(* IEC 61131-3 sources: OpenPlc_Lezioni/Blocchi_PorteLogiche/build, 2 files *)

(* ---- plc.st ---- *)
TYPE
  LOGLEVEL : (CRITICAL, WARNING, INFO, DEBUG) := INFO;
END_TYPE

FUNCTION_BLOCK LOGGER
  VAR_INPUT
    TRIG : BOOL;
    MSG : STRING;
    LEVEL : LOGLEVEL := INFO;
  END_VAR
  VAR
    TRIG0 : BOOL;
  END_VAR

  IF TRIG AND NOT TRIG0 THEN
  {{
   LogMessage(GetFbVar(LEVEL),(char*)GetFbVar(MSG, .body),GetFbVar(MSG, .len));
  }}
  END_IF;
  TRIG0:=TRIG;
END_FUNCTION_BLOCK

PROGRAM program0
  VAR
    P1 : BOOL;
    P2 : BOOL;
    P3 : BOOL;
    P4 : BOOL;
    P5 : BOOL;
    P6 : BOOL;
    P7 : BOOL;
    LED1 : BOOL;
    LED2 : BOOL;
    LED3 : BOOL;
    LED4 : BOOL;
    _TMP_AND1_OUT : BOOL;
    _TMP_OR2_OUT : BOOL;
    _TMP_AND10_OUT : BOOL;
    _TMP_NOT18_OUT : BOOL;
  END_VAR

  _TMP_AND1_OUT := AND(P1, P2);
  LED1 := _TMP_AND1_OUT;
  _TMP_OR2_OUT := OR(P3, P4);
  LED2 := _TMP_OR2_OUT;
  _TMP_AND10_OUT := AND(P5, P6);
  LED2 := _TMP_AND10_OUT;
  _TMP_NOT18_OUT := NOT(P7);
  LED4 := _TMP_NOT18_OUT;
END_PROGRAM

CONFIGURATION Config0

  RESOURCE Res0 ON PLC
    TASK task0(INTERVAL := T#20ms,PRIORITY := 0);
    PROGRAM instance0 WITH task0 : program0;
  END_RESOURCE
END_CONFIGURATION

(* ---- generated_plc.st ---- *)
PROGRAM program0
  VAR
    P1 : BOOL;
    P2 : BOOL;
    P3 : BOOL;
    P4 : BOOL;
    P5 : BOOL;
    P6 : BOOL;
    P7 : BOOL;
    LED1 : BOOL;
    LED2 : BOOL;
    LED3 : BOOL;
    LED4 : BOOL;
    _TMP_AND1_OUT : BOOL;
    _TMP_OR2_OUT : BOOL;
    _TMP_AND10_OUT : BOOL;
    _TMP_NOT18_OUT : BOOL;
  END_VAR

  _TMP_AND1_OUT := AND(P1, P2);
  LED1 := _TMP_AND1_OUT;
  _TMP_OR2_OUT := OR(P3, P4);
  LED2 := _TMP_OR2_OUT;
  _TMP_AND10_OUT := AND(P5, P6);
  LED2 := _TMP_AND10_OUT;
  _TMP_NOT18_OUT := NOT(P7);
  LED4 := _TMP_NOT18_OUT;
END_PROGRAM

CONFIGURATION Config0

  RESOURCE Res0 ON PLC
    TASK task0(INTERVAL := T#20ms,PRIORITY := 0);
    PROGRAM instance0 WITH task0 : program0;
  END_RESOURCE
END_CONFIGURATION
